Fanuc KAREL source: kb00127.compact.KL

PROGRAM KB00127
%STACKSIZE=65535
%PRIORITY=65535
%NOLOCKGROUP
VAR
P1 : STRING[80]
P2 : INTEGER
RESULT : INTEGER
BEGIN
P1='A'
P2=1
RESULT=ORD(P1,P2)
END KB00127
